{region 'Documentation'}
(*!
<summary>Check that IN is at most Maximum.</summary>
<description>

All checked operands and bounds must be finite; NaN or either infinity reports Error
during active evaluation.

Numeric diagnostics use the formatter's default six significant digits; rounding affects
the message only, not the comparison.

</description>
*)
{endregion}
FUNCTION_BLOCK AssertLessEqual_Real EXTENDS AssertionBase
VAR_INPUT
    IN : REAL; //! Actual value checked or observed by this Assertion.
    Maximum : REAL; //! Inclusive upper bound of the comparison; for a range, must not be below Minimum.
END_VAR

SUPER^();

{region 'Documentation'}
(*!
<summary>Check that IN is at most Maximum.</summary>
*)
{endregion}
METHOD PROTECTED Assert
VAR
    Message : STRING(GVL_Constants.MessageLength);
    MaximumText : STRING(GVL_Constants.AssertionValueLength);
    ActualText : STRING(GVL_Constants.AssertionValueLength);
END_VAR
IF NOT EvaluationActive THEN
    RETURN;
END_IF;

IF Result = E_Result.Error THEN
    RETURN;
END_IF;

IF NOT Tc2_Utilities.RealIsFinite(x := IN) THEN
    Error(Message := 'Assertion error: IN must be finite.');
    RETURN;
END_IF;

IF NOT Tc2_Utilities.RealIsFinite(x := Maximum) THEN
    Error(Message := 'Assertion error: Maximum must be finite.');
    RETURN;
END_IF;

IF Result = E_Result.Failed THEN
    RETURN;
END_IF;

IF IN > Maximum THEN
    MaximumText := CreateAssertionTextValue_Real(Value := Maximum);
    ActualText := CreateAssertionTextValue_Real(Value := IN);
    Message := CONCAT('Assertion failed: value is above maximum. Maximum = ',
        MaximumText);
    Message := CONCAT(Message, ', Actual = ');
    Message := CONCAT(Message, ActualText);
    Message := CONCAT(Message, '.');
    Fail(Message := Message);
    RETURN;
END_IF;

Pass();
END_METHOD

END_FUNCTION_BLOCK

(* stored: Version 1.1.0.1
   POU AssertLessEqual_Real: Id {4df76200-1677-4439-be10-c9c01ba13091}, SpecialFunc None
   Folder Internal: Id {2b3960bc-5d38-4e3b-ae42-55178cc929a9}
   Method Assert: Id {6bed8024-8c98-43c7-ab6d-7ddbd7b026ce} *)
